Staubli VAL3: utBorder.pjx

--- utBorder.pjx ---
Parameters version=s8.8.3Cs9_BS1660 stackSize=5000 millimeterUnit=true
Program file=start.pgx
Program file=stop.pgx
Data file=utBorder.dtx

--- utBorder.dtx ---
public string sBorderColour

--- start.pgx ---
program start()
begin
end

--- stop.pgx ---
program stop()
begin
end
